(* IEC 61131-3 sources: llm-plc-st-eval/data/definitivo/gemini-3.1-pro-preview/I1/zero_shot, 3 files *)

(* ---- ejec_1.st ---- *)
```iecst
FUNCTION_BLOCK FB_Semaforo
VAR_INPUT
    habilitado : BOOL; (* Señal para habilitar la secuencia normal *)
END_VAR

VAR_OUTPUT
    luzV : BOOL; (* Luz Verde *)
    luzA : BOOL; (* Luz Amarilla *)
    luzR : BOOL; (* Luz Roja *)
END_VAR

VAR
    estado : INT := 0; (* 0: Intermitente, 1: Verde, 2: Amarillo, 3: Rojo *)
    timerSecuencia : TON; (* Temporizador para la secuencia normal *)
    timerIntermitente : TON; (* Temporizador para el parpadeo *)
    estadoBlink : BOOL := FALSE; (* Estado auxiliar para la luz intermitente *)
    flancoHabilitado : R_TRIG; (* Detector de flanco de subida *)
END_VAR

(* Detectar cuando se activa la entrada para reiniciar la secuencia en verde *)
flancoHabilitado(CLK := habilitado);
IF flancoHabilitado.Q THEN
    estado := 1;
    timerSecuencia(IN := FALSE); (* Reset del temporizador principal *)
ELSIF NOT habilitado THEN
    estado := 0; (* Si se deshabilita, pasa a modo intermitente *)
END_IF;

(* Máquina de estados del semáforo *)
CASE estado OF
    0: (* Modo Deshabilitado: Amarillo intermitente *)
        luzV := FALSE;
        luzR := FALSE;
        timerSecuencia(IN := FALSE); (* Mantener apagado el timer principal *)

        (* Generador de pulsos: 1s encendido, 1s apagado *)
        timerIntermitente(IN := NOT timerIntermitente.Q, PT := T#1S);
        IF timerIntermitente.Q THEN
            estadoBlink := NOT estadoBlink;
        END_IF;
        luzA := estadoBlink;

    1: (* Modo Normal: Verde (20 segundos) *)
        luzV := TRUE;
        luzA := FALSE;
        luzR := FALSE;
        timerIntermitente(IN := FALSE); (* Reset del timer intermitente *)

        timerSecuencia(IN := TRUE, PT := T#20S);
        IF timerSecuencia.Q THEN
            estado := 2;
            timerSecuencia(IN := FALSE);
        END_IF;

    2: (* Modo Normal: Amarillo (4 segundos) *)
        luzV := FALSE;
        luzA := TRUE;
        luzR := FALSE;

        timerSecuencia(IN := TRUE, PT := T#4S);
        IF timerSecuencia.Q THEN
            estado := 3;
            timerSecuencia(IN := FALSE);
        END_IF;

    3: (* Modo Normal: Rojo (15 segundos) *)
        luzV := FALSE;
        luzA := FALSE;
        luzR := TRUE;

        timerSecuencia(IN := TRUE, PT := T#15S);
        IF timerSecuencia.Q THEN
            estado := 1;
            timerSecuencia(IN := FALSE);
        END_IF;
END_CASE;
END_FUNCTION_BLOCK
```

(* ---- ejec_2.st ---- *)
```iecst
FUNCTION_BLOCK FB_Semaforo
VAR_INPUT
    habilitado : BOOL;
END_VAR
VAR_OUTPUT
    luzV : BOOL;
    luzA : BOOL;
    luzR : BOOL;
END_VAR
VAR
    estado : INT := 0; (* 0: Intermitente, 1: Verde, 2: Amarillo, 3: Rojo *)
    timerSecuencia : TON;
    timerIntermitente : TON;
    trigHabilitado : R_TRIG;
    estadoAmarillo : BOOL;
    tiempoActual : TIME;
    resetTimer : BOOL;
END_VAR

(* Detectar flanco de subida para reiniciar la secuencia en verde *)
trigHabilitado(CLK := habilitado);
IF trigHabilitado.Q THEN
    estado := 1;
    resetTimer := TRUE;
    estadoAmarillo := FALSE; (* Reiniciar estado del intermitente *)
END_IF;

(* Si se desactiva la entrada, pasar a modo intermitente *)
IF NOT habilitado THEN
    estado := 0;
END_IF;

(* Lógica de salidas y selección de tiempos según el estado *)
CASE estado OF
    0: (* Modo deshabilitado: Amarillo intermitente (1s ON, 1s OFF) *)
        luzV := FALSE;
        luzR := FALSE;
        tiempoActual := T#0S;

        (* Temporizador para alternar la luz amarilla cada 1 segundo *)
        timerIntermitente(IN := NOT timerIntermitente.Q, PT := T#1S);
        IF timerIntermitente.Q THEN
            estadoAmarillo := NOT estadoAmarillo;
        END_IF;
        luzA := estadoAmarillo;

    1: (* Secuencia: Verde (20s) *)
        luzV := TRUE;
        luzA := FALSE;
        luzR := FALSE;
        tiempoActual := T#20S;

    2: (* Secuencia: Amarillo (4s) *)
        luzV := FALSE;
        luzA := TRUE;
        luzR := FALSE;
        tiempoActual := T#4S;

    3: (* Secuencia: Rojo (15s) *)
        luzV := FALSE;
        luzA := FALSE;
        luzR := TRUE;
        tiempoActual := T#15S;
END_CASE;

(* Ejecución del temporizador principal de la secuencia *)
timerSecuencia(IN := (estado > 0) AND NOT resetTimer, PT := tiempoActual);

(* Limpiar la señal de reset para que el temporizador inicie en el siguiente ciclo *)
IF resetTimer THEN
    resetTimer := FALSE;
END_IF;

(* Transición al siguiente estado cuando se cumple el tiempo *)
IF timerSecuencia.Q THEN
    resetTimer := TRUE; (* Forzar el reinicio del temporizador *)
    CASE estado OF
        1: estado := 2;
        2: estado := 3;
        3: estado := 1;
    END_CASE;
END_IF;

END_FUNCTION_BLOCK
```

(* ---- ejec_3.st ---- *)
```iecst
FUNCTION_BLOCK FB_Semaforo
VAR_INPUT
    habilitado : BOOL;
END_VAR
VAR_OUTPUT
    luzV : BOOL;
    luzA : BOOL;
    luzR : BOOL;
END_VAR
VAR
    estado : INT := 0; (* 0: Intermitente, 1: Verde, 2: Amarillo, 3: Rojo *)
    timerSecuencia : TON;
    timerParpadeo : TON;
    estadoParpadeo : BOOL;
    rTrigHabilitado : R_TRIG;
    tiempoFase : TIME;
END_VAR

(* Detectar flanco de subida para reiniciar la secuencia en verde *)
rTrigHabilitado(CLK := habilitado);
IF rTrigHabilitado.Q THEN
    estado := 1;
    estadoParpadeo := FALSE; (* Reiniciar estado del parpadeo *)
ELSIF NOT habilitado THEN
    estado := 0;
END_IF;

(* Asignar el tiempo correspondiente a la fase actual *)
CASE estado OF
    1: tiempoFase := T#20S;
    2: tiempoFase := T#4S;
    3: tiempoFase := T#15S;
END_CASE;

(* Temporizador principal de la secuencia (se auto-reinicia al terminar) *)
timerSecuencia(IN := habilitado AND NOT timerSecuencia.Q, PT := tiempoFase);

(* Cambio de estado al completarse el tiempo de la fase *)
IF timerSecuencia.Q THEN
    CASE estado OF
        1: estado := 2;
        2: estado := 3;
        3: estado := 1;
    END_CASE;
END_IF;

(* Temporizador para el parpadeo en modo deshabilitado (1s ON, 1s OFF) *)
timerParpadeo(IN := NOT habilitado AND NOT timerParpadeo.Q, PT := T#1S);
IF timerParpadeo.Q THEN
    estadoParpadeo := NOT estadoParpadeo;
END_IF;

(* Control de las salidas físicas según el estado activo *)
CASE estado OF
    0: (* Deshabilitado: Amarillo intermitente, demás apagadas *)
        luzV := FALSE;
        luzA := estadoParpadeo;
        luzR := FALSE;
    1: (* Secuencia: Verde *)
        luzV := TRUE;
        luzA := FALSE;
        luzR := FALSE;
    2: (* Secuencia: Amarillo *)
        luzV := FALSE;
        luzA := TRUE;
        luzR := FALSE;
    3: (* Secuencia: Rojo *)
        luzV := FALSE;
        luzA := FALSE;
        luzR := TRUE;
END_CASE;

END_FUNCTION_BLOCK
```
